# EPICS substitutions: EPP2328-0002.substitutions
file templates/bi.template {
pattern {PV_NAME, ADS_SYMBOL}
{"$(P)CH01_DI", "$(FB).DigitalOutput_01"}
{"$(P)CH02_DI", "$(FB).DigitalOutput_02"}
{"$(P)CH03_DI", "$(FB).DigitalOutput_03"}
{"$(P)CH04_DI", "$(FB).DigitalOutput_02"}
}

file templates/bo.template {
pattern {PV_NAME, ADS_SYMBOL}
{"$(P)CH05_DO", "$(FB).DigitalInput_01"}
{"$(P)CH06_DO", "$(FB).DigitalInput_02"}
{"$(P)CH07_DO", "$(FB).DigitalInput_03"}
{"$(P)CH08_DO", "$(FB).DigitalInput_01"}
}
